// TIA Portal V21 program export: 0 tag tables, 0 data types, 0 data blocks, 2 code blocks (in call order from the OBs), 0 instance data blocks

ORGANIZATION_BLOCK "CallAndCompare"   // OB1, LAD
   VAR_TEMP   // added for the SCL form of the ladder/FBD networks
      _w1 : Bool;
   END_VAR
BEGIN

REGION Network 1: Pump on high level
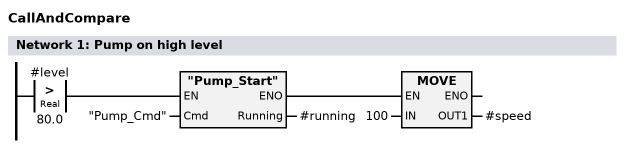
   RUNG wire#powerrail
      { S7_Templates := "SrcType := Real" } GT_Contact(in1 := #level, in2 := 80.0)
      "Pump_Start"(Cmd := "Pump_Cmd", Running => #running)
      Move(in := 100, out1 => #speed)
   END_RUNG
   // the same network as SCL:
   "Pump_Start"(EN := #level > 80.0, Cmd := "Pump_Cmd", Running => #running, ENO => #_w1);
   IF #_w1 THEN #speed := 100; END_IF;
END_REGION
END_ORGANIZATION_BLOCK

FUNCTION_BLOCK "Mixed"   // FB1, LAD
BEGIN

REGION Network 1: Unknown part
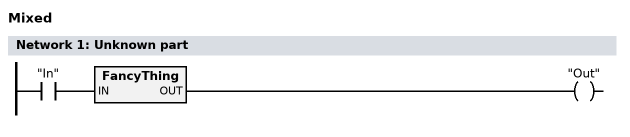
   // no SCL statement known for FancyThing: written as a call
   "Out" := FancyThing("In");
END_REGION

REGION Network 2 (SCL): SCL inside
END_REGION

REGION Network 3: Empty
END_REGION
END_FUNCTION_BLOCK
